# EPICS substitutions: db/Beckhoff_7XXX/ecmcEL7411_OPT_inputs.substitutions
file "ecmcEL7411_OPT_inputs.template"
{
  pattern {CH_ID}
          {"$(OPT_CH_ID=01)"}
}
